// TIA Portal V20 export
TYPE "Stoermeldung"
   STRUCT
      SM : Array[0..127] of Bool;
   END_STRUCT;
END_TYPE
